(* IEC 61131-3 sources: kns-port-domestic/tools/port_metrics_tests/fixtures/adapted/src/POUs/PRG_Main, 1 file *)

(* ---- PRG_Main.decl.st ---- *)
PROGRAM PRG_Main
VAR
    fbPump : FB_Pump;
    xStartCmd : BOOL;
    xSimulation : BOOL; // PORT: [foo] режим имитации
END_VAR
